ABB RAPID module: SubProg.mod

MODULE MOD_SubProg

PERS wobjdata rdkWObj := [FALSE, TRUE, "", [[0,0,0],[1,0,0,0]],[[0,0,0],[1,0,0,0]]];
PERS tooldata rdkTool := [TRUE,[[0,0,0],[1,0,0,0]],[6.8,[0,0,15],[1,0,0,0],0,0,0.005]];
VAR speeddata rdkSpeed := [500,500,500,500];
VAR zonedata rdkZone := z1;
VAR extjoint rdkExtax := [9E9,9E9,9E9,9E9,9E9,9E9];

PROC main_RoboDK()
	SubProg;
	EXIT;
ENDPROC

PROC SubProg()
	!Program generated by RoboDK v5.9.4 for ABB IRB 1600-8/1.45 on 26/10/2026 01:01:07
	!Using nominal kinematics.
	var robtarget crt;
	crt := CRobT(\Tool:=rdkTool, \WObj:=rdkWObj);
	rdkExtax := crt.extax;
	ConfJ \On;
	ConfL \Off;
	rdkWObj.uframe:=[[0.000,0.000,0.000],[1.00000000,0.00000000,0.00000000,0.00000000]];
	rdkWObj.oframe:=[[851.624,-621.056,1118.740],[0.96592583,0.00000000,0.00000000,0.25881905]];
	rdkTool.tframe:=[[0.000,0.000,120.000],[0.99144486,0.00000000,0.13052619,0.00000001]];
	MoveL [[0.000,0.000,0.000],[0.58801837,0.20533497,0.76632048,-0.15755906],[-1,-1,0,1],rdkExtax], rdkSpeed, rdkZone, rdkTool, \WObj:=rdkWObj;
	!Inside sub
ENDPROC

ENDMODULE
